(*
SPDX-FileCopyrightText: © 2026 Oleksandr Tiutyk <trofimich@gmail.com>
SPDX-License-Identifier: MIT
License: https://opensource.org/license/mit
*)

(*!
<summary>Groups workflow ownership, topology, configuration, failure handling and timing scenarios.</summary>
<description>Owns the fixed case tree and runs its leaves in order in the controller task.</description>
*)

{attribute 'no_assign'}
{attribute 'no_explicit_call' := 'do not call this function block directly'}
FUNCTION_BLOCK WorkflowContractTestGroup EXTENDS TOF_Testing.TestGroup<28>
VAR_STAT
	{attribute 'hide'}
	_ClassName : STRING := __POUNAME();
END_VAR
VAR
	_RootAssociation : WorkflowContractTestCase(
		name := "TestRootAssociation",
		parent := THIS^,
		scenario := WORKFLOW_CONTRACT_TEST_SCENARIO.ROOT_ASSOCIATION
	);
	_SequenceTopology : WorkflowContractTestCase(
		name := "TestSequenceTopology",
		parent := THIS^,
		scenario := WORKFLOW_CONTRACT_TEST_SCENARIO.SEQUENCE_TOPOLOGY
	);
	_TransitionDiagnostics : WorkflowContractTestCase(
		name := "TestTransitionDiagnostics",
		parent := THIS^,
		scenario := WORKFLOW_CONTRACT_TEST_SCENARIO.TRANSITION_DIAGNOSTICS
	);
	_DependencyBindings : WorkflowContractTestCase(
		name := "TestDependencyBindings",
		parent := THIS^,
		scenario := WORKFLOW_CONTRACT_TEST_SCENARIO.DEPENDENCY_BINDINGS
	);
	_WriteConfiguration : WorkflowContractTestCase(
		name := "TestWriteConfiguration",
		parent := THIS^,
		scenario := WORKFLOW_CONTRACT_TEST_SCENARIO.WRITE_CONFIGURATION
	);
	_LoadConfiguration : WorkflowContractTestCase(
		name := "TestLoadConfiguration",
		parent := THIS^,
		scenario := WORKFLOW_CONTRACT_TEST_SCENARIO.LOAD_CONFIGURATION
	);
	_OperatorSerialization : WorkflowContractTestCase(
		name := "TestOperatorSerialization",
		parent := THIS^,
		scenario := WORKFLOW_CONTRACT_TEST_SCENARIO.OPERATOR_SERIALIZATION
	);
	_DeserializeNullContextRejection : WorkflowContractTestCase(
		name := "TestDeserializeNullContextRejection",
		parent := THIS^,
		scenario := WORKFLOW_CONTRACT_TEST_SCENARIO.DESERIALIZE_NULL_CONTEXT_REJECTION
	);
	_FactoryDeclarations : WorkflowContractTestCase(
		name := "TestFactoryDeclarations",
		parent := THIS^,
		scenario := WORKFLOW_CONTRACT_TEST_SCENARIO.FACTORY_DECLARATIONS
	);
	_ArrayValidation : WorkflowContractTestCase(
		name := "TestArrayValidation",
		parent := THIS^,
		scenario := WORKFLOW_CONTRACT_TEST_SCENARIO.ARRAY_VALIDATION
	);
	_WorkflowIsolation : WorkflowContractTestCase(
		name := "TestWorkflowIsolation",
		parent := THIS^,
		scenario := WORKFLOW_CONTRACT_TEST_SCENARIO.WORKFLOW_ISOLATION
	);
	_ConditionTopology : WorkflowContractTestCase(
		name := "TestConditionTopology",
		parent := THIS^,
		scenario := WORKFLOW_CONTRACT_TEST_SCENARIO.CONDITION_TOPOLOGY
	);
	_ParentSetters : WorkflowContractTestCase(
		name := "TestParentSetters",
		parent := THIS^,
		scenario := WORKFLOW_CONTRACT_TEST_SCENARIO.PARENT_SETTERS
	);
	_InitializationRetry : WorkflowContractTestCase(
		name := "TestInitializationRetry",
		parent := THIS^,
		scenario := WORKFLOW_CONTRACT_TEST_SCENARIO.INITIALIZATION_RETRY
	);
	_BoundaryDiagnostics : WorkflowContractTestCase(
		name := "TestBoundaryDiagnostics",
		parent := THIS^,
		scenario := WORKFLOW_CONTRACT_TEST_SCENARIO.BOUNDARY_DIAGNOSTICS
	);
	_InvokeConfiguration : WorkflowContractTestCase(
		name := "TestInvokeConfiguration",
		parent := THIS^,
		scenario := WORKFLOW_CONTRACT_TEST_SCENARIO.INVOKE_CONFIGURATION
	);
	_TaskFailureDuringSuspend : WorkflowContractTestCase(
		name := "TestTaskFailureDuringSuspend",
		parent := THIS^,
		scenario := WORKFLOW_CONTRACT_TEST_SCENARIO.TASK_FAILURE_DURING_SUSPEND
	);
	_TaskCompletionDuringSuspend : WorkflowContractTestCase(
		name := "TestTaskCompletionDuringSuspend",
		parent := THIS^,
		scenario := WORKFLOW_CONTRACT_TEST_SCENARIO.TASK_COMPLETION_DURING_SUSPEND
	);
	_TaskAbortDuringSuspend : WorkflowContractTestCase(
		name := "TestTaskAbortDuringSuspend",
		parent := THIS^,
		scenario := WORKFLOW_CONTRACT_TEST_SCENARIO.TASK_ABORT_DURING_SUSPEND
	);
	_TaskReleaseFailureDuringCancel : WorkflowContractTestCase(
		name := "TestTaskReleaseFailureDuringCancel",
		parent := THIS^,
		scenario := WORKFLOW_CONTRACT_TEST_SCENARIO.TASK_RELEASE_FAILURE_DURING_CANCEL
	);
	_CatchCleanupBoundary : WorkflowContractTestCase(
		name := "TestCatchCleanupBoundary",
		parent := THIS^,
		scenario := WORKFLOW_CONTRACT_TEST_SCENARIO.CATCH_CLEANUP_BOUNDARY
	);
	_ConcreteMetadata : WorkflowContractTestCase(
		name := "TestConcreteMetadata",
		parent := THIS^,
		scenario := WORKFLOW_CONTRACT_TEST_SCENARIO.CONCRETE_METADATA
	);
	_VariableLookup : WorkflowContractTestCase(
		name := "TestVariableLookup",
		parent := THIS^,
		scenario := WORKFLOW_CONTRACT_TEST_SCENARIO.VARIABLE_LOOKUP
	);
	_DeclaredVariableReset : WorkflowContractTestCase(
		name := "TestDeclaredVariableReset",
		parent := THIS^,
		scenario := WORKFLOW_CONTRACT_TEST_SCENARIO.DECLARED_VARIABLE_RESET
	);
	_DeclaredVariableValidation : WorkflowContractTestCase(
		name := "TestDeclaredVariableValidation",
		parent := THIS^,
		scenario := WORKFLOW_CONTRACT_TEST_SCENARIO.DECLARED_VARIABLE_VALIDATION
	);
	_ConditionScopePrecedence : WorkflowContractTestCase(
		name := "TestConditionScopePrecedence",
		parent := THIS^,
		scenario := WORKFLOW_CONTRACT_TEST_SCENARIO.CONDITION_SCOPE_PRECEDENCE
	);
	_DelayPauseRemaining : WorkflowDelayPauseRemainingTest(name := "TestDelayPauseRemaining", parent := THIS^);
	_DelayLifecycle : WorkflowContractTestCase(
		name := "TestDelayLifecycle",
		parent := THIS^,
		scenario := WORKFLOW_CONTRACT_TEST_SCENARIO.DELAY_LIFECYCLE
	);
END_VAR
VAR
	_Children : ARRAY [0.._ChildCount - 1] OF TOF_Testing.ITestElement :=
	[
		_RootAssociation,
		_SequenceTopology,
		_TransitionDiagnostics,
		_DependencyBindings,
		_WriteConfiguration,
		_LoadConfiguration,
		_OperatorSerialization,
		_DeserializeNullContextRejection,
		_FactoryDeclarations,
		_ArrayValidation,
		_WorkflowIsolation,
		_ConditionTopology,
		_ParentSetters,
		_InitializationRetry,
		_BoundaryDiagnostics,
		_InvokeConfiguration,
		_TaskFailureDuringSuspend,
		_TaskCompletionDuringSuspend,
		_TaskAbortDuringSuspend,
		_TaskReleaseFailureDuringCancel,
		_CatchCleanupBoundary,
		_ConcreteMetadata,
		_VariableLookup,
		_DeclaredVariableReset,
		_DeclaredVariableValidation,
		_ConditionScopePrecedence,
		_DelayPauseRemaining,
		_DelayLifecycle
	];
END_VAR

(*!
<summary>Borrows the persistent case array. Callers must not modify it.</summary>
*)
{attribute 'monitoring' := 'call'}
PROPERTY Children : REFERENCE TO ARRAY [0.._ChildCount - 1] OF TOF_Testing.ITestElement
GET
Children REF= _Children;
END_GET
END_PROPERTY

(*!
<summary>Borrows the concrete class name. Callers must not modify it.</summary>
*)
{attribute 'monitoring' := 'call'}
PROPERTY ClassName : REFERENCE TO STRING
GET
ClassName REF= _ClassName;
END_GET
END_PROPERTY

(*!
<summary>Borrows the project namespace name. Callers must not modify it.</summary>
*)
{attribute 'monitoring' := 'call'}
PROPERTY NamespaceName : REFERENCE TO STRING
GET
NamespaceName REF= CurrentNamespace.Name;
END_GET
END_PROPERTY

(*!
<summary>Reports the complete instance size in bytes.</summary>
*)
{attribute 'monitoring' := 'call'}
PROPERTY SelfSize : ULINT
GET
SelfSize := XSIZEOF(THIS^);
END_GET
END_PROPERTY

END_FUNCTION_BLOCK

(* stored: Version 1.1.0.1
   POU WorkflowContractTestGroup: Id {a9fd8154-d63b-4fcf-af02-d6981feca319}, SpecialFunc None
   Property Children: Id {bcceda25-6b85-41a2-9533-d767f4461eea}
   Get Get: Id {f9f53561-fb7b-4fd4-89c3-bd74ffe63987}
   Property ClassName: Id {22e4f8c0-473d-40f7-ba6c-1ce62e365cc4}
   Get Get: Id {e29809bc-3fb3-4545-9d52-c3894e252a62}
   Property NamespaceName: Id {15b5521e-489e-4f3b-810d-6ef38dab3423}
   Get Get: Id {5df929c9-b285-4cc5-9d2a-91646bdd085a}
   Property SelfSize: Id {65bbafa7-977f-437a-bf1b-d3f124fbd5b1}
   Get Get: Id {01222d6b-14dc-4eae-8741-83d199d1d80f} *)
